(* IEC 61131-3 sources: yaads/test/twincat/plc, 8 files *)

(* ---- E_Mode.st ---- *)
// DUT E_Mode
{attribute 'qualified_only'}
TYPE E_Mode :
(
    eOff := 0,
    eAuto := 1,
    eManual := 2
) INT;
END_TYPE

(* ---- ST_Flags.st ---- *)
// DUT ST_Flags: two BITs in the first byte, and a BYTE after them
TYPE ST_Flags :
STRUCT
    bA    : BIT;
    bB    : BIT;
    nRest : BYTE;
END_STRUCT
END_TYPE

(* ---- ST_Packed.st ---- *)
// DUT ST_Packed: no padding at all
{attribute 'pack_mode' := '1'}
TYPE ST_Packed :
STRUCT
    nSmall : SINT;
    fBig   : LREAL;
END_STRUCT
END_TYPE

(* ---- ST_Pump.st ---- *)
// DUT ST_Pump: laid out by TwinCAT 3's default pack_mode, 8
TYPE ST_Pump :
STRUCT
    nSpeed   : INT;
    fTemp    : LREAL;
    bRunning : BOOL;
    eMode    : E_Mode;
    sTag     : STRING(10);
END_STRUCT
END_TYPE

(* ---- U_Value.st ---- *)
// DUT U_Value
TYPE U_Value :
UNION
    nDint  : DINT;
    fReal  : REAL;
    aBytes : ARRAY [0..3] OF BYTE;
END_UNION
END_TYPE

(* ---- GVL.st ---- *)
// GVL GVL
VAR_GLOBAL
    {attribute 'TcEncoding' := 'UTF-8'}
    sUtf8 : STRING(20);
END_VAR

(* ---- GVL_Long.st ---- *)
// GVL GVL_Long: the 64-bit dates and times, from TwinCAT 3.1.4026 on; leave it out before that
VAR_GLOBAL
    ldDate   : LDATE;
    ldtStamp : LDATE_AND_TIME;
    ltodTime : LTIME_OF_DAY;
END_VAR

(* ---- MAIN.st ---- *)
// POU MAIN, a PROGRAM in Structured Text, called by the PLC task
PROGRAM MAIN
VAR
    // as ADS.Test.FakePLC has them
    nCounter : DINT;
    nSpeed   : INT;
    bOn      : BOOL;
    fTemp    : LREAL;
    sName    : STRING(20);
    wsText   : WSTRING(10);
    aValues  : ARRAY [1..5] OF INT;
    stPump   : ST_Pump;
    aPumps   : ARRAY [0..1] OF ST_Pump;
    eMode    : E_Mode;
    tDelay   : TIME;
    dtStamp  : DATE_AND_TIME;
    sText    : T_MaxString;
    stFlags  : ST_Flags;

    // the rest of the elementary types
    nSint    : SINT;
    nUsint   : USINT;
    nUint    : UINT;
    nUdint   : UDINT;
    nLint    : LINT;
    nUlint   : ULINT;
    nByte    : BYTE;
    nWord    : WORD;
    nDword   : DWORD;
    nLword   : LWORD;
    fReal    : REAL;
    tLong    : LTIME;
    dDate    : DATE;
    todTime  : TIME_OF_DAY;

    // and of the others
    aMatrix  : ARRAY [0..1, -1..1] OF INT;
    stPacked : ST_Packed;
    uValue   : U_Value;
    pnSpeed  : POINTER TO INT;
    aBig     : ARRAY [0..599] OF USINT;

    // counts the cycles, for the cyclic notifications
    nTicks   : UDINT;
END_VAR

nTicks := nTicks + 1;
pnSpeed := ADR(nSpeed);
